// Mitsubishi GX Works2 project: mqttrobotplc   PLC: Q03UDV

PROGRAM MAIN
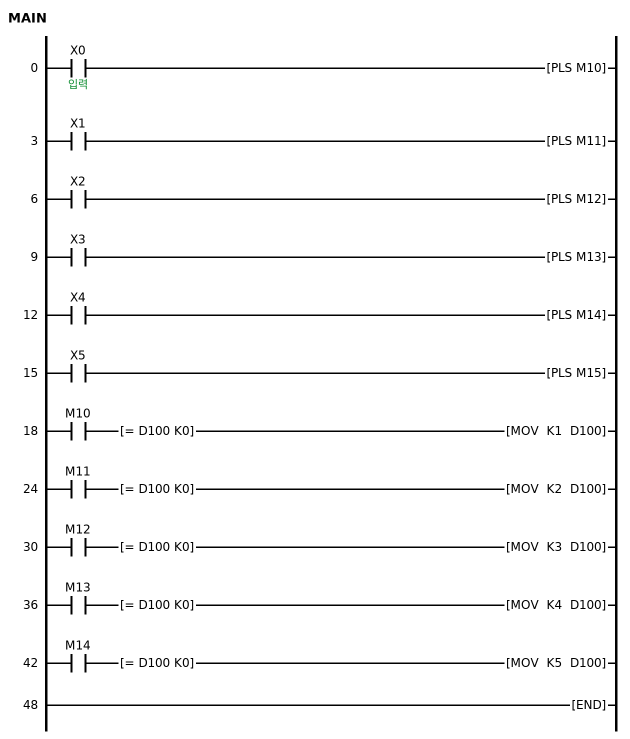
0     LD      X0  ; 입력
      PLS     M10
3     LD      X1
      PLS     M11
6     LD      X2
      PLS     M12
9     LD      X3
      PLS     M13
12    LD      X4
      PLS     M14
15    LD      X5
      PLS     M15
18    LD      M10
      AND=    D100 K0
      MOV     K1 D100
24    LD      M11
      AND=    D100 K0
      MOV     K2 D100
30    LD      M12
      AND=    D100 K0
      MOV     K3 D100
36    LD      M13
      AND=    D100 K0
      MOV     K4 D100
42    LD      M14
      AND=    D100 K0
      MOV     K5 D100
48    END
END_PROGRAM
